(* IEC 61131-3 sources: SafePLC-Gen-Evaluation/Evaluation Results/dexpi/run_04, 2 files *)

(* ---- io_declarations.st ---- *)
(* ==================================================  *)
(* PLC I/O Variable Declarations — CODESYS 3.5  *)
(* Generated by SafePLC-Gen Multimodal  *)
(* ==================================================  *)

VAR_GLOBAL
    (* --- Analog Inputs ---  *)
    PI_4712.01_Raw               AT %IW0       : INT := 0;    (* PI-4712.01 — Pressure indicator (local gauge) on disc  *)
    PICSA_4712.02_Raw            AT %IW2       : INT := 0;    (* PICSA-4712.02 — Pressure indicator, controller, switch w  *)
    TICSA_4750.03_Raw            AT %IW4       : INT := 0;    (* TICSA-4750.03 — Temperature indicator, controller, switc  *)
    (* --- Analog Outputs ---  *)
    PV_4712.02_Out               AT %QW0       : INT := 0;    (* PV-4712.02 — Pressure control valve, fail-closed (F.C  *)
    TV_4750.03_Out               AT %QW2       : INT := 0;    (* TV-4750.03 — Temperature control valve, fail-open (F.  *)
    (* --- Digital Inputs ---  *)
    HS_4750.01                   AT %IX0.0     : BOOL := FALSE;    (* HS-4750.01 — Hand switch (operator pushbutton or sele  *)
    (* --- Digital Outputs ---  *)
    XV_4750.01                   AT %QX0.0     : BOOL := FALSE;    (* XV-4750.01 — Solenoid-operated on/off valve, fail-clo  *)
END_VAR

(* ---- generated_code.st ---- *)
(* Generated by SafePLC-Gen Multimodal — CODESYS 3.5 *)
(* IEC 61131-3 Structured Text *)
(* Date: 2026-04-25T11:49:41.344215 *)

PROGRAM PLC_PRG

VAR
    TICSA_4750_03_Raw            AT %IW4       : INT := 0;
    PICSA_4712_02_Raw            AT %IW2       : INT := 0;
    PI_4712_01_Raw               AT %IW0       : INT := 0;
    HS_4750_01                   AT %IX0.0     : BOOL := FALSE;
    TV_4750_03_Out               AT %QW2       : INT := 0;
    PV_4712_02_Out               AT %QW0       : INT := 0;
    XV_4750_01                   AT %QX0.0     : BOOL := FALSE;
    ESTOP                        AT %IX0.1     : BOOL := FALSE;
    MANUAL_RESET                 AT %IX0.2     : BOOL := FALSE;
END_VAR

VAR
    FirstScan                    : BOOL := TRUE;

    TICSA_4750_03_Scaled         : REAL := 0.0;
    PICSA_4712_02_Scaled         : REAL := 0.0;
    PI_4712_01_Scaled            : REAL := 0.0;

    TICSA_4750_03_SP             : REAL := 80.0;
    TICSA_4750_03_HH_SP          : REAL := 110.0;
    TICSA_4750_03_H_SP           : REAL := 100.0;
    TICSA_4750_03_L_SP           : REAL := 20.0;
    TICSA_4750_03_LL_SP          : REAL := 10.0;
    TICSA_4750_03_Deadband       : REAL := 2.0;
    TICSA_4750_03_H              : BOOL := FALSE;
    TICSA_4750_03_L              : BOOL := FALSE;
    TICSA_4750_03_HH_Latch       : SR := (S1 := FALSE, R := FALSE, Q1 := FALSE);
    TICSA_4750_03_LL_Latch       : SR := (S1 := FALSE, R := FALSE, Q1 := FALSE);
    TICSA_4750_03_HH_Ack         : BOOL := FALSE;
    TICSA_4750_03_LL_Ack         : BOOL := FALSE;

    PICSA_4712_02_SP             : REAL := 5.0;
    PICSA_4712_02_HH_SP          : REAL := 9.0;
    PICSA_4712_02_H_SP           : REAL := 8.0;
    PICSA_4712_02_L_SP           : REAL := 1.0;
    PICSA_4712_02_LL_SP          : REAL := 0.5;
    PICSA_4712_02_Deadband       : REAL := 0.2;
    PICSA_4712_02_H              : BOOL := FALSE;
    PICSA_4712_02_L              : BOOL := FALSE;
    PICSA_4712_02_HH_Latch       : SR := (S1 := FALSE, R := FALSE, Q1 := FALSE);
    PICSA_4712_02_LL_Latch       : SR := (S1 := FALSE, R := FALSE, Q1 := FALSE);
    PICSA_4712_02_HH_Ack         : BOOL := FALSE;
    PICSA_4712_02_LL_Ack         : BOOL := FALSE;

    PI_4712_01_HH_SP             : REAL := 9.5;
    PI_4712_01_H_SP              : REAL := 8.5;
    PI_4712_01_L_SP              : REAL := 0.8;
    PI_4712_01_LL_SP             : REAL := 0.3;
    PI_4712_01_Deadband          : REAL := 0.2;
    PI_4712_01_H                 : BOOL := FALSE;
    PI_4712_01_L                 : BOOL := FALSE;
    PI_4712_01_HH_Latch          : SR := (S1 := FALSE, R := FALSE, Q1 := FALSE);
    PI_4712_01_LL_Latch          : SR := (S1 := FALSE, R := FALSE, Q1 := FALSE);
    PI_4712_01_HH_Ack            : BOOL := FALSE;
    PI_4712_01_LL_Ack            : BOOL := FALSE;

    LOOP_4750_03_TRIP            : BOOL := FALSE;
    LOOP_4712_02_TRIP            : BOOL := FALSE;
    LOOP_104_01_TRIP             : BOOL := FALSE;
    TICSA_4750_03_HH             : BOOL := FALSE;
    TICSA_4750_03_LL             : BOOL := FALSE;
    PICSA_4712_02_HH             : BOOL := FALSE;
    PICSA_4712_02_LL             : BOOL := FALSE;
    SV_104_01_HH                 : BOOL := FALSE;
    SV_104_01_LL                 : BOOL := FALSE;
    SAFE_STATE                   : BOOL := FALSE;

    TIC_Error                    : REAL := 0.0;
    TIC_Integral                 : REAL := 0.0;
    TIC_Kp                       : REAL := 1.2;
    TIC_Ki                       : REAL := 0.05;
    TIC_Output                   : REAL := 0.0;

    PIC_Error                    : REAL := 0.0;
    PIC_Integral                 : REAL := 0.0;
    PIC_Kp                       : REAL := 1.5;
    PIC_Ki                       : REAL := 0.08;
    PIC_Output                   : REAL := 0.0;

    SV_104_01_Out                : BOOL := FALSE;
    HV_MNb_47123_ISO_Out         : BOOL := FALSE;
    CHK_73KH12_50_P4712_Out      : BOOL := FALSE;
    CHK_MNc_47124_P4712_Out      : BOOL := FALSE;
    STR_75SA21_80_Out            : BOOL := FALSE;
    BV_75HB13_73HG12_Out         : BOOL := FALSE;
    BV_Q_80_N6_Out               : BOOL := FALSE;
    HV_QSa_47140_Out             : BOOL := FALSE;
    HV_QSb_47141_Out             : BOOL := FALSE;
    SB_Q_80_N6_Out               : BOOL := FALSE;

    System_Alarm                 : BOOL := FALSE;
END_VAR

IF FirstScan THEN
    LOOP_4750_03_TRIP := TRUE;
    LOOP_4712_02_TRIP := TRUE;
    LOOP_104_01_TRIP  := TRUE;
    SAFE_STATE        := TRUE;
    TV_4750_03_Out    := 32767;
    PV_4712_02_Out    := 6554;
    XV_4750_01        := FALSE;
    SV_104_01_Out              := FALSE;
    HV_MNb_47123_ISO_Out       := FALSE;
    CHK_73KH12_50_P4712_Out    := FALSE;
    CHK_MNc_47124_P4712_Out    := FALSE;
    STR_75SA21_80_Out          := FALSE;
    BV_75HB13_73HG12_Out       := FALSE;
    BV_Q_80_N6_Out             := FALSE;
    HV_QSa_47140_Out           := FALSE;
    HV_QSb_47141_Out           := FALSE;
    SB_Q_80_N6_Out             := FALSE;
    FirstScan         := FALSE;
    RETURN;
END_IF;

TICSA_4750_03_Scaled := ((INT_TO_REAL(TICSA_4750_03_Raw) - 6554.0) / (32767.0 - 6554.0)) * 150.0;
PICSA_4712_02_Scaled := ((INT_TO_REAL(PICSA_4712_02_Raw) - 6554.0) / (32767.0 - 6554.0)) * 10.0;
PI_4712_01_Scaled    := ((INT_TO_REAL(PI_4712_01_Raw)    - 6554.0) / (32767.0 - 6554.0)) * 10.0;

TICSA_4750_03_HH := TICSA_4750_03_Scaled > TICSA_4750_03_HH_SP;
TICSA_4750_03_LL := TICSA_4750_03_Scaled < TICSA_4750_03_LL_SP;
PICSA_4712_02_HH := PICSA_4712_02_Scaled > PICSA_4712_02_HH_SP;
PICSA_4712_02_LL := PICSA_4712_02_Scaled < PICSA_4712_02_LL_SP;
SV_104_01_HH     := HS_4750_01;
SV_104_01_LL     := FALSE;

IF TICSA_4750_03_HH OR TICSA_4750_03_LL THEN
    LOOP_4750_03_TRIP := TRUE;
ELSIF LOOP_4750_03_TRIP AND MANUAL_RESET
      AND NOT TICSA_4750_03_HH AND NOT TICSA_4750_03_LL THEN
    LOOP_4750_03_TRIP := FALSE;
END_IF;

IF PICSA_4712_02_HH OR PICSA_4712_02_LL THEN
    LOOP_4712_02_TRIP := TRUE;
ELSIF LOOP_4712_02_TRIP AND MANUAL_RESET
      AND NOT PICSA_4712_02_HH AND NOT PICSA_4712_02_LL THEN
    LOOP_4712_02_TRIP := FALSE;
END_IF;

IF SV_104_01_HH OR SV_104_01_LL THEN
    LOOP_104_01_TRIP := TRUE;
ELSIF LOOP_104_01_TRIP AND MANUAL_RESET
      AND NOT SV_104_01_HH AND NOT SV_104_01_LL THEN
    LOOP_104_01_TRIP := FALSE;
END_IF;

SAFE_STATE := ESTOP
              OR LOOP_4750_03_TRIP
              OR LOOP_4712_02_TRIP
              OR LOOP_104_01_TRIP;

IF NOT SAFE_STATE THEN
    TIC_Error    := TICSA_4750_03_SP - TICSA_4750_03_Scaled;
    TIC_Integral := TIC_Integral + (TIC_Ki * TIC_Error);
    IF TIC_Integral > 100.0 THEN
        TIC_Integral := 100.0;
    ELSIF TIC_Integral < 0.0 THEN
        TIC_Integral := 0.0;
    END_IF;
    TIC_Output := (TIC_Kp * TIC_Error) + TIC_Integral;
    IF TIC_Output > 100.0 THEN
        TIC_Output := 100.0;
    ELSIF TIC_Output < 0.0 THEN
        TIC_Output := 0.0;
    END_IF;
    TV_4750_03_Out := REAL_TO_INT(6554.0 + (TIC_Output / 100.0) * (32767.0 - 6554.0));
ELSE
    TV_4750_03_Out := 32767;
END_IF;

IF NOT SAFE_STATE THEN
    PIC_Error    := PICSA_4712_02_SP - PICSA_4712_02_Scaled;
    PIC_Integral := PIC_Integral + (PIC_Ki * PIC_Error);
    IF PIC_Integral > 100.0 THEN
        PIC_Integral := 100.0;
    ELSIF PIC_Integral < 0.0 THEN
        PIC_Integral := 0.0;
    END_IF;
    PIC_Output := (PIC_Kp * PIC_Error) + PIC_Integral;
    IF PIC_Output > 100.0 THEN
        PIC_Output := 100.0;
    ELSIF PIC_Output < 0.0 THEN
        PIC_Output := 0.0;
    END_IF;
    PV_4712_02_Out := REAL_TO_INT(6554.0 + (PIC_Output / 100.0) * (32767.0 - 6554.0));
ELSE
    PV_4712_02_Out := 6554;
END_IF;

IF NOT SAFE_STATE AND HS_4750_01 THEN
    XV_4750_01 := TRUE;
ELSE
    XV_4750_01 := FALSE;
END_IF;

IF NOT SAFE_STATE THEN
    SV_104_01_Out            := TRUE;
    HV_MNb_47123_ISO_Out     := TRUE;
    CHK_73KH12_50_P4712_Out  := TRUE;
    CHK_MNc_47124_P4712_Out  := TRUE;
    STR_75SA21_80_Out        := TRUE;
    BV_75HB13_73HG12_Out     := TRUE;
    BV_Q_80_N6_Out           := TRUE;
    HV_QSa_47140_Out         := TRUE;
    HV_QSb_47141_Out         := TRUE;
    SB_Q_80_N6_Out           := TRUE;
ELSE
    SV_104_01_Out            := FALSE;
    HV_MNb_47123_ISO_Out     := FALSE;
    CHK_73KH12_50_P4712_Out  := FALSE;
    CHK_MNc_47124_P4712_Out  := FALSE;
    STR_75SA21_80_Out        := FALSE;
    BV_75HB13_73HG12_Out     := FALSE;
    BV_Q_80_N6_Out           := FALSE;
    HV_QSa_47140_Out         := FALSE;
    HV_QSb_47141_Out         := FALSE;
    SB_Q_80_N6_Out           := FALSE;
END_IF;

(* Four-level alarms — TICSA-4750.03 *)
IF TICSA_4750_03_Scaled > TICSA_4750_03_HH_SP THEN
    TICSA_4750_03_HH_Latch.S1 := TRUE;
ELSIF TICSA_4750_03_Scaled <= (TICSA_4750_03_HH_SP - TICSA_4750_03_Deadband) THEN
    TICSA_4750_03_HH_Latch.S1 := FALSE;
END_IF;
TICSA_4750_03_HH_Latch.R := TICSA_4750_03_HH_Ack AND NOT TICSA_4750_03_HH;
TICSA_4750_03_HH_Latch(S1 := TICSA_4750_03_HH_Latch.S1, R := TICSA_4750_03_HH_Latch.R);

IF TICSA_4750_03_Scaled > TICSA_4750_03_H_SP THEN
    TICSA_4750_03_H := TRUE;
ELSIF TICSA_4750_03_Scaled <= (TICSA_4750_03_H_SP - TICSA_4750_03_Deadband) THEN
    TICSA_4750_03_H := FALSE;
END_IF;

IF TICSA_4750_03_Scaled < TICSA_4750_03_L_SP THEN
    TICSA_4750_03_L := TRUE;
ELSIF TICSA_4750_03_Scaled >= (TICSA_4750_03_L_SP + TICSA_4750_03_Deadband) THEN
    TICSA_4750_03_L := FALSE;
END_IF;

IF TICSA_4750_03_Scaled < TICSA_4750_03_LL_SP THEN
    TICSA_4750_03_LL_Latch.S1 := TRUE;
ELSIF TICSA_4750_03_Scaled >= (TICSA_4750_03_LL_SP + TICSA_4750_03_Deadband) THEN
    TICSA_4750_03_LL_Latch.S1 := FALSE;
END_IF;
TICSA_4750_03_LL_Latch.R := TICSA_4750_03_LL_Ack AND NOT TICSA_4750_03_LL;
TICSA_4750_03_LL_Latch(S1 := TICSA_4750_03_LL_Latch.S1, R := TICSA_4750_03_LL_Latch.R);

(* Four-level alarms — PICSA-4712.02 *)
IF PICSA_4712_02_Scaled > PICSA_4712_02_HH_SP THEN
    PICSA_4712_02_HH_Latch.S1 := TRUE;
ELSIF PICSA_4712_02_Scaled <= (PICSA_4712_02_HH_SP - PICSA_4712_02_Deadband) THEN
    PICSA_4712_02_HH_Latch.S1 := FALSE;
END_IF;
PICSA_4712_02_HH_Latch.R := PICSA_4712_02_HH_Ack AND NOT PICSA_4712_02_HH;
PICSA_4712_02_HH_Latch(S1 := PICSA_4712_02_HH_Latch.S1, R := PICSA_4712_02_HH_Latch.R);

IF PICSA_4712_02_Scaled > PICSA_4712_02_H_SP THEN
    PICSA_4712_02_H := TRUE;
ELSIF PICSA_4712_02_Scaled <= (PICSA_4712_02_H_SP - PICSA_4712_02_Deadband) THEN
    PICSA_4712_02_H := FALSE;
END_IF;

IF PICSA_4712_02_Scaled < PICSA_4712_02_L_SP THEN
    PICSA_4712_02_L := TRUE;
ELSIF PICSA_4712_02_Scaled >= (PICSA_4712_02_L_SP + PICSA_4712_02_Deadband) THEN
    PICSA_4712_02_L := FALSE;
END_IF;

IF PICSA_4712_02_Scaled < PICSA_4712_02_LL_SP THEN
    PICSA_4712_02_LL_Latch.S1 := TRUE;
ELSIF PICSA_4712_02_Scaled >= (PICSA_4712_02_LL_SP + PICSA_4712_02_Deadband) THEN
    PICSA_4712_02_LL_Latch.S1 := FALSE;
END_IF;
PICSA_4712_02_LL_Latch.R := PICSA_4712_02_LL_Ack AND NOT PICSA_4712_02_LL;
PICSA_4712_02_LL_Latch(S1 := PICSA_4712_02_LL_Latch.S1, R := PICSA_4712_02_LL_Latch.R);

(* Four-level alarms — PI-4712.01 *)
IF PI_4712_01_Scaled > PI_4712_01_HH_SP THEN
    PI_4712_01_HH_Latch.S1 := TRUE;
ELSIF PI_4712_01_Scaled <= (PI_4712_01_HH_SP - PI_4712_01_Deadband) THEN
    PI_4712_01_HH_Latch.S1 := FALSE;
END_IF;
PI_4712_01_HH_Latch.R := PI_4712_01_HH_Ack AND NOT (PI_4712_01_Scaled > PI_4712_01_HH_SP);
PI_4712_01_HH_Latch(S1 := PI_4712_01_HH_Latch.S1, R := PI_4712_01_HH_Latch.R);

IF PI_4712_01_Scaled > PI_4712_01_H_SP THEN
    PI_4712_01_H := TRUE;
ELSIF PI_4712_01_Scaled <= (PI_4712_01_H_SP - PI_4712_01_Deadband) THEN
    PI_4712_01_H := FALSE;
END_IF;

IF PI_4712_01_Scaled < PI_4712_01_L_SP THEN
    PI_4712_01_L := TRUE;
ELSIF PI_4712_01_Scaled >= (PI_4712_01_L_SP + PI_4712_01_Deadband) THEN
    PI_4712_01_L := FALSE;
END_IF;

IF PI_4712_01_Scaled < PI_4712_01_LL_SP THEN
    PI_4712_01_LL_Latch.S1 := TRUE;
ELSIF PI_4712_01_Scaled >= (PI_4712_01_LL_SP + PI_4712_01_Deadband) THEN
    PI_4712_01_LL_Latch.S1 := FALSE;
END_IF;
PI_4712_01_LL_Latch.R := PI_4712_01_LL_Ack AND NOT (PI_4712_01_Scaled < PI_4712_01_LL_SP);
PI_4712_01_LL_Latch(S1 := PI_4712_01_LL_Latch.S1, R := PI_4712_01_LL_Latch.R);

System_Alarm :=
    TICSA_4750_03_HH_Latch.Q1 OR TICSA_4750_03_LL_Latch.Q1 OR
    TICSA_4750_03_H            OR TICSA_4750_03_L            OR
    PICSA_4712_02_HH_Latch.Q1 OR PICSA_4712_02_LL_Latch.Q1 OR
    PICSA_4712_02_H            OR PICSA_4712_02_L            OR
    PI_4712_01_HH_Latch.Q1    OR PI_4712_01_LL_Latch.Q1    OR
    PI_4712_01_H               OR PI_4712_01_L               OR
    LOOP_4750_03_TRIP          OR LOOP_4712_02_TRIP          OR
    LOOP_104_01_TRIP           OR SAFE_STATE;

END_PROGRAM
